            ELSIF fbReceive.nRecBytes > 0 THEN
                nRxCount := nRxCount + fbReceive.nRecBytes;
                IF nRxCount >= 9 THEN
                    nExpectedFrame := 9 + BYTE_TO_UDINT(aRx[7]) + BYTE_TO_UDINT(aRx[8]) * 256;
                    IF (nExpectedFrame < 11) OR (nExpectedFrame > SIZEOF(aRx)) THEN
                        bError := TRUE; nErrorID := 16#E104;
                        stSession.bConnected := FALSE;
                        bBusy := FALSE; nState := 0;
                    ELSIF nRxCount >= nExpectedFrame THEN
                        IF (aRx[0] <> 16#D0) OR (aRx[1] <> 16#00) THEN
                            bError := TRUE; nErrorID := 16#E105;
                            stSession.bConnected := FALSE;
                        ELSE
                            nEndCode := BYTE_TO_UINT(aRx[9]) + BYTE_TO_UINT(aRx[10]) * 256;
                            IF nEndCode <> 0 THEN
                                bError := TRUE; nErrorID := nEndCode;
                            ELSIF (bBitAccess AND (nExpectedFrame < 11 + ((UINT_TO_UDINT(nPoints) + 1) / 2)))
                                 OR ((NOT bBitAccess) AND (nExpectedFrame < 11 + UINT_TO_UDINT(nPoints) * 2)) THEN
                                bError := TRUE; nErrorID := 16#E107;
                                stSession.bConnected := FALSE;
                            ELSE
                                IF bBitAccess THEN
                                    pDestBit := pData;
                                    FOR nIdx := 0 TO (UINT_TO_UDINT(nPoints) - 1) DO
                                        IF (nIdx MOD 2) = 0 THEN
                                            pDestBit[nIdx] := ((aRx[11 + (nIdx / 2)] AND 16#10) <> 0);
                                        ELSE
                                            pDestBit[nIdx] := ((aRx[11 + (nIdx / 2)] AND 16#01) <> 0);
                                        END_IF;
                                    END_FOR;
                                ELSE
                                    pDestByte := pData;
                                    nCopyBytes := UINT_TO_UDINT(nPoints) * 2;
                                    FOR nIdx := 0 TO (nCopyBytes - 1) DO
                                        pDestByte[nIdx] := aRx[11 + nIdx];
                                    END_FOR;
                                END_IF;
                                bDone := TRUE;
                            END_IF;
                        END_IF;
                        bBusy := FALSE; nState := 0;
                    ELSE
                        nState := 20; // Fragment received; wait for rest of frame
                    END_IF;
                ELSE
                    nState := 20; // Header itself is fragmented
                END_IF;

            ELSIF tonTimeout.Q THEN
                // Quá 2 giây không có phản hồi
                bError   := TRUE;
                nErrorID := 16#E103; // Timeout chờ response
                stSession.bConnected := FALSE;
                bBusy    := FALSE;
                nState   := 0;

            ELSE
                // Chưa có dữ liệu về trong scan này -> Kích đọc tiếp ở scan sau
                nState := 20;
            END_IF;
        END_IF;

END_CASE;

// Cập nhật trạng thái bận vào session dùng chung
// Only the FB that acquired the socket lock may release it.
IF bBusy THEN
    stSession.bBusy := TRUE;
ELSIF bOwnsSession THEN
    stSession.bBusy := FALSE;
    bOwnsSession := FALSE;
END_IF;

END_FUNCTION_BLOCK

// ---- POUs/FB_MelsecDebugXY4Pt.TcPOU
FUNCTION_BLOCK FB_MelsecDebugXY4Pt
VAR_INPUT
    bExecute          : BOOL := FALSE; // Rising edge for ONE 4-point DATA-ONLY test
    bPermit           : BOOL := FALSE; // Maintenance gate, OFF by default
    bMachineStopped   : BOOL := FALSE; // Axis, encoder and gantry are stationary
    bPublisherIdle    : BOOL := FALSE; // All live motion publishers inhibited
    bAbort            : BOOL := FALSE; // Cancel the data-only sequence
    rCenterX_mm       : LREAL := 50.0;
    rCenterY_mm       : LREAL := 85.0;
    rAngleDeg         : LREAL := 0.0;
    rLength_mm        : LREAL := 40.0;
    rWidth_mm         : LREAL := 40.0;
    tHold             : TIME := T#10S; // GX Works2 observation pause, NOT motion acknowledgment
END_VAR
VAR_IN_OUT
    stSession         : ST_MelsecSession; // Same owned socket as all other TwinCAT FBs
END_VAR
VAR_OUTPUT
    bBusy             : BOOL;
    bDone             : BOOL;       // Four XY frames READ BACK; NOT robot motion completion
    bError            : BOOL;
    nErrorCode        : INT;
    nCommErrorID      : UDINT;
    nState            : INT := 0;
    nCurrentVertex    : INT;        // 1..4, stays at 4 after success
    nPassedVertices   : INT;
    nWriteX           : DINT;
    nWriteY           : DINT;
    nReadX            : DINT;
    nReadY            : DINT;
    nReadVertex       : UINT;
    bLastReadbackOK   : BOOL;
    bAllMotionBitsLow : BOOL;
    bOriginalRestored : BOOL; // Original XY/index restored after all four hold windows
END_VAR
VAR
    fbStart           : R_TRIG;
    fbWrite           : FB_MelsecWrite;
    fbRead            : FB_MelsecRead;
    tonHold           : TON;
    aCorners          : ARRAY[1..4] OF ST_Point2D;
    rAngleRad         : LREAL;
    rC                : LREAL;
    rS                : LREAL;
    rHL               : LREAL;
    rHW               : LREAL;
    aXYWrite          : ARRAY[0..1] OF DINT;
    aXYRead           : ARRAY[0..1] OF DINT;
    nIndexWrite       : UINT;
    nIndexRead        : UINT;
    aOriginalXY       : ARRAY[0..1] OF DINT;
    nOriginalIndex    : UINT;
    bNeedSnapshot     : BOOL;
    bRestoring        : BOOL;
    aStartAck         : ARRAY[0..1] OF BOOL; // M1000 M1001
    aRobotFlags       : ARRAY[0..3] OF BOOL; // M102, M103, M104, M105
    nPlcFsmState      : DINT;               // D200/D201
    bWriteReq         : BOOL;
    bReadReq          : BOOL;
    eReadDevice       : E_MelsecDevice;
    nReadAddress      : UDINT;
    nReadPoints       : UINT;
    bReadBitMode      : BOOL;
    pReadData         : PVOID;
    nReadDataSize     : UDINT;
    nWriteAddress     : UDINT;
    nWritePoints      : UINT;
    pWriteData        : PVOID;
    nWriteDataSize    : UDINT;
END_VAR

// Diagnostic mode NEVER writes M1000 or any PLC bit, never touches Z.
// Only D100..D103 (2x DINT XY) and D114 (UINT vertex) are ever written.
// Explicit machine-stopped conditions are checked on EVERY scan.
fbStart(CLK := bExecute);
tonHold(IN := (nState = 20), PT := tHold);

bReadReq := FALSE;
bWriteReq := FALSE;

IF (nState <> 0) AND (nState <> 99) AND (NOT bPermit OR NOT bMachineStopped OR
    NOT bPublisherIdle OR bAbort OR NOT stSession.bConnected) THEN
    bError := TRUE;
    nErrorCode := 901; // Lost permit, motion interlock, or TCP
    nState := 99;
END_IF;

CASE nState OF
    0: // IDLE - no automatic restart
        bBusy := FALSE;
        IF fbStart.Q THEN
            bDone := FALSE;
            bError := FALSE;
            bLastReadbackOK := FALSE;
            bAllMotionBitsLow := FALSE;
            nPassedVertices := 0;
            nCurrentVertex := 0;
            bNeedSnapshot := TRUE;
            bRestoring := FALSE;
            bOriginalRestored := FALSE;
            nErrorCode := 0;
            nCommErrorID := 0;
            IF NOT bPermit OR NOT bMachineStopped OR NOT bPublisherIdle
                OR bAbort OR NOT stSession.bConnected OR stSession.bBusy THEN
                bError := TRUE; nErrorCode := 901;
            ELSIF (rLength_mm <= 0.0) OR (rWidth_mm <= 0.0)
                OR (rLength_mm > 100.0) OR (rWidth_mm > 100.0)
                OR (tHold < T#2S) OR (tHold > T#60S) THEN
                bError := TRUE; nErrorCode := 902;
            ELSE
                rAngleRad := rAngleDeg * 3.141592653589793 / 180.0;
                rC := COS(rAngleRad);
                rS := SIN(rAngleRad);
                rHL := rLength_mm / 2.0;
                rHW := rWidth_mm / 2.0;

                aCorners[1].X := rCenterX_mm + rHL * rC - rHW * rS;
                aCorners[1].Y := rCenterY_mm + rHL * rS + rHW * rC;
                aCorners[2].X := rCenterX_mm - rHL * rC - rHW * rS;
                aCorners[2].Y := rCenterY_mm - rHL * rS + rHW * rC;
                aCorners[3].X := rCenterX_mm - rHL * rC + rHW * rS;
                aCorners[3].Y := rCenterY_mm - rHL * rS - rHW * rC;
                aCorners[4].X := rCenterX_mm + rHL * rC + rHW * rS;
                aCorners[4].Y := rCenterY_mm + rHL * rS - rHW * rC;

                nCurrentVertex := 1;
                bBusy := TRUE;
                nState := 1;
            END_IF;
        END_IF;

    // Recheck Mitsubishi handshake before EVERY vertex (read-only).
    1:
        eReadDevice := DEV_M; nReadAddress := 1000; nReadPoints := 2;
        bReadBitMode := TRUE;
        pReadData := ADR(aStartAck); nReadDataSize := SIZEOF(aStartAck);
        bReadReq := TRUE;
        nState := 2;

    2:
        IF fbRead.bDone THEN
            IF aStartAck[0] OR aStartAck[1] THEN
                bError := TRUE; nErrorCode := 903; nState := 99;
            ELSE
                nState := 3;
            END_IF;
        ELSIF fbRead.bError THEN
            bError := TRUE; nErrorCode := 910; nCommErrorID := fbRead.nErrorID; nState := 99;
        END_IF;

    3:
        eReadDevice := DEV_M; nReadAddress := 102; nReadPoints := 4;
        bReadBitMode := TRUE;
        pReadData := ADR(aRobotFlags); nReadDataSize := SIZEOF(aRobotFlags);
        bReadReq := TRUE;
        nState := 4;

    4:
        IF fbRead.bDone THEN
            IF aRobotFlags[0] OR aRobotFlags[1] OR aRobotFlags[2] OR aRobotFlags[3] THEN
                bError := TRUE; nErrorCode := 904; nState := 99;
            ELSE
                nState := 5;
            END_IF;
        ELSIF fbRead.bError THEN
            bError := TRUE; nErrorCode := 911; nCommErrorID := fbRead.nErrorID; nState := 99;
        END_IF;

    5:
        eReadDevice := DEV_D; nReadAddress := 200; nReadPoints := 2;
        bReadBitMode := FALSE;
        pReadData := ADR(nPlcFsmState); nReadDataSize := SIZEOF(nPlcFsmState);
        bReadReq := TRUE;
        nState := 6;

    6:
        IF fbRead.bDone THEN
            IF nPlcFsmState <> 0 THEN
                bError := TRUE; nErrorCode := 905; nState := 99;
            ELSE
                bAllMotionBitsLow := TRUE;
                IF bRestoring THEN
                    nState := 30;
                ELSIF bNeedSnapshot THEN
                    nState := 7;
                ELSE
                    nState := 10;
                END_IF;
            END_IF;
        ELSIF fbRead.bError THEN
            bError := TRUE; nErrorCode := 912; nCommErrorID := fbRead.nErrorID; nState := 99;
        END_IF;

    7: // Snapshot original XY before any data-only write
        eReadDevice := DEV_D; nReadAddress := 100; nReadPoints := 4;
        bReadBitMode := FALSE;
        pReadData := ADR(aOriginalXY); nReadDataSize := SIZEOF(aOriginalXY);
        bReadReq := TRUE;
        nState := 8;

    8:
        IF fbRead.bDone THEN
            nState := 9;
        ELSIF fbRead.bError THEN
            bError := TRUE; nErrorCode := 918; nCommErrorID := fbRead.nErrorID; nState := 99;
        END_IF;

    9:
        eReadDevice := DEV_D; nReadAddress := 114; nReadPoints := 1;
        bReadBitMode := FALSE;
        pReadData := ADR(nOriginalIndex); nReadDataSize := SIZEOF(nOriginalIndex);
        bReadReq := TRUE;
        nState := 91;

    91:
        IF fbRead.bDone THEN
            bNeedSnapshot := FALSE;
            nState := 10;
        ELSIF fbRead.bError THEN
            bError := TRUE; nErrorCode := 919; nCommErrorID := fbRead.nErrorID; nState := 99;
        END_IF;

    10: // Data-only: two DINTs. Deliberately no Z/speed write.
        IF (nCurrentVertex < 1) OR (nCurrentVertex > 4) OR
            (aCorners[nCurrentVertex].X < 5.0) OR
            (aCorners[nCurrentVertex].X > 170.0) OR
            (aCorners[nCurrentVertex].Y < 5.0) OR
            (aCorners[nCurrentVertex].Y > 165.0) THEN
            bError := TRUE; nErrorCode := 906; nState := 99;
        ELSE
            nWriteX := LREAL_TO_DINT(aCorners[nCurrentVertex].X * 10000.0);
            nWriteY := LREAL_TO_DINT(aCorners[nCurrentVertex].Y * 10000.0);
            aXYWrite[0] := nWriteX;
            aXYWrite[1] := nWriteY;
            nIndexWrite := INT_TO_UINT(nCurrentVertex);
            nWriteAddress := 100; nWritePoints := 4;
            pWriteData := ADR(aXYWrite); nWriteDataSize := SIZEOF(aXYWrite);
            bLastReadbackOK := FALSE;
            bWriteReq := TRUE;
            nState := 11;
        END_IF;

    11:
        IF fbWrite.bDone THEN
            nState := 12;
        ELSIF fbWrite.bError THEN
            bError := TRUE; nErrorCode := 913; nCommErrorID := fbWrite.nErrorID; nState := 99;
        END_IF;

    12: // Different rising edge for D114
        nWriteAddress := 114; nWritePoints := 1;
        pWriteData := ADR(nIndexWrite); nWriteDataSize := SIZEOF(nIndexWrite);
        bWriteReq := TRUE;
        nState := 13;

    13:
        IF fbWrite.bDone THEN
            nState := 14;
        ELSIF fbWrite.bError THEN
            bError := TRUE; nErrorCode := 914; nCommErrorID := fbWrite.nErrorID; nState := 99;
        END_IF;

    14:
        eReadDevice := DEV_D; nReadAddress := 100; nReadPoints := 4;
        bReadBitMode := FALSE;
        pReadData := ADR(aXYRead); nReadDataSize := SIZEOF(aXYRead);
        bReadReq := TRUE;
        nState := 15;

    15:
        IF fbRead.bDone THEN
            nState := 16;
        ELSIF fbRead.bError THEN
            bError := TRUE; nErrorCode := 915; nCommErrorID := fbRead.nErrorID; nState := 99;
        END_IF;

    16:
        eReadDevice := DEV_D; nReadAddress := 114; nReadPoints := 1;
        bReadBitMode := FALSE;
        pReadData := ADR(nIndexRead); nReadDataSize := SIZEOF(nIndexRead);
        bReadReq := TRUE;
        nState := 17;

    17:
        IF fbRead.bDone THEN
            nReadX := aXYRead[0];
            nReadY := aXYRead[1];
            nReadVertex := nIndexRead;
            bLastReadbackOK := (nReadX = nWriteX) AND (nReadY = nWriteY)
                               AND (nReadVertex = nIndexWrite);
            IF bLastReadbackOK THEN
                nPassedVertices := nPassedVertices + 1;
                nState := 20; // Hold for operator GX Works2 observation
            ELSE
                bError := TRUE; nErrorCode := 916; nState := 99;
            END_IF;
        ELSIF fbRead.bError THEN
            bError := TRUE; nErrorCode := 917; nCommErrorID := fbRead.nErrorID; nState := 99;
        END_IF;

    20: // Observation timer. Never mislabel elapsed time as QD75 motion ACK.
        IF tonHold.Q THEN
            IF nCurrentVertex >= 4 THEN
                bRestoring := TRUE;
                bAllMotionBitsLow := FALSE;
                nState := 1; // Recheck M1000/ACK/BUSY/FSM before restoring original packet
            ELSE
                nCurrentVertex := nCurrentVertex + 1;
                bAllMotionBitsLow := FALSE;
                nState := 1;
            END_IF;
        END_IF;

    30: // Restore original XY, then original index: never leave stale debug target
        nWriteAddress := 100; nWritePoints := 4;
        pWriteData := ADR(aOriginalXY); nWriteDataSize := SIZEOF(aOriginalXY);
        bWriteReq := TRUE;
        nState := 31;

    31:
        IF fbWrite.bDone THEN
            nState := 32;
        ELSIF fbWrite.bError THEN
            bError := TRUE; nErrorCode := 920; nCommErrorID := fbWrite.nErrorID; nState := 99;
        END_IF;

    32:
        nWriteAddress := 114; nWritePoints := 1;
        pWriteData := ADR(nOriginalIndex); nWriteDataSize := SIZEOF(nOriginalIndex);
        bWriteReq := TRUE;
        nState := 33;

    33:
        IF fbWrite.bDone THEN
            nState := 34;
        ELSIF fbWrite.bError THEN
            bError := TRUE; nErrorCode := 921; nCommErrorID := fbWrite.nErrorID; nState := 99;
        END_IF;

    34:
        eReadDevice := DEV_D; nReadAddress := 100; nReadPoints := 4;
        bReadBitMode := FALSE;
        pReadData := ADR(aXYRead); nReadDataSize := SIZEOF(aXYRead);
        bReadReq := TRUE;
        nState := 35;

    35:
        IF fbRead.bDone THEN
            nState := 36;
        ELSIF fbRead.bError THEN
            bError := TRUE; nErrorCode := 922; nCommErrorID := fbRead.nErrorID; nState := 99;
        END_IF;

    36:
        eReadDevice := DEV_D; nReadAddress := 114; nReadPoints := 1;
        bReadBitMode := FALSE;
        pReadData := ADR(nIndexRead); nReadDataSize := SIZEOF(nIndexRead);
        bReadReq := TRUE;
        nState := 37;

    37:
        IF fbRead.bDone THEN
            bOriginalRestored := (aXYRead[0] = aOriginalXY[0]) AND
                (aXYRead[1] = aOriginalXY[1]) AND (nIndexRead = nOriginalIndex);
            IF bOriginalRestored THEN
                bBusy := FALSE;
                bDone := TRUE; // All 4 readbacks AND full restore confirmed
                nState := 0;
            ELSE
                bError := TRUE; nErrorCode := 923; nState := 99;
            END_IF;
        ELSIF fbRead.bError THEN
            bError := TRUE; nErrorCode := 924; nCommErrorID := fbRead.nErrorID; nState := 99;
        END_IF;

    99: // Latched diagnostic failure. NO reset command sent to the PLC.
        bBusy := FALSE;
        bDone := FALSE;
        bReadReq := FALSE;
        bWriteReq := FALSE;
        IF NOT bExecute AND NOT bPermit AND NOT fbRead.bBusy AND NOT fbWrite.bBusy THEN
            nState := 0;
        END_IF;
END_CASE;

// READS may access only M1000,M1001,M102..M105,D200..D201,D100..D103,D114.
// WRITES are strictly limited to D100..D103 and D114, never M, Z or QD75.
fbWrite(
    stSession := stSession, bExecute := bWriteReq,
    eDevice := DEV_D, nStartAddr := nWriteAddress,
    nPoints := nWritePoints, bBitAccess := FALSE,
    pData := pWriteData, nDataSize := nWriteDataSize
);
fbRead(
    stSession := stSession, bExecute := bReadReq,
    eDevice := eReadDevice, nStartAddr := nReadAddress,
    nPoints := nReadPoints, bBitAccess := bReadBitMode,
    pData := pReadData, nDataSize := nReadDataSize
);

END_FUNCTION_BLOCK

// ---- POUs/FB_UpstreamCameraTracking4Pt.TcPOU
FUNCTION_BLOCK FB_UpstreamCameraTracking4Pt
VAR_INPUT
    bReset               : BOOL;
    bCameraResult        : BOOL;  // Single rising edge: camera provides center and angle ONLY
    bAcceptCamera        : BOOL;
    bCalibrationConfirmed: BOOL;  // NEVER assume Camera and Robot coordinates coincide
    bExposureEncoderValid : BOOL; // Capture encoder synchronized with IMAGE EXPOSURE, not processing result
    rEncoderAtExposure_mm : LREAL; // Encoder latched by TwinCAT when camera takes the image
    rCameraCenterX_mm    : LREAL; // Already calibrated from pixels into millimeters
    rCameraCenterY_mm    : LREAL;
    rCameraAngleDeg      : LREAL;
    rCameraToWorkStart_mm : LREAL; // USER INPUT after calibration: Camera trigger station to ROBOT X=0, positive mm
    rCameraToRobotX_mm   : LREAL; // Fine X calibration correction only; NOT the Camera->Robot distance
    rCameraToRobotY_mm   : LREAL;
    rCameraToRobotYawDeg : LREAL; // Calibrated camera-to-robot axis angle
    rEncoderTotalDist_mm : LREAL; // Continuous integrated encoder distance, not 16-bit count
    rLength_mm           : LREAL := 40.0;
    rWidth_mm            : LREAL := 40.0;
    rRobotXMin_mm        : LREAL := 0.0;
    rRobotXMax_mm        : LREAL := 180.0;
    rRobotYMin_mm        : LREAL := 0.0;
    rRobotYMax_mm        : LREAL := 170.0;
END_VAR
VAR_OUTPUT
    bCaptured            : BOOL; // Product retained while travelling FROM camera to robot
    bInRobotWorkspace    : BOOL; // At least one corner in workspace (diagnostic only)
    bAllCornersPastRobot : BOOL;
    bCalibrationMissing  : BOOL;
    nCaptureCount        : UDINT;
    nRejectedCount       : UDINT;
    nErrorCode           : INT;
    rEncoderAtCapture_mm : LREAL;
    rEncoderTravel_mm    : LREAL;
    rCenterAtCaptureX_mm : LREAL; // Robot reference frame at camera trigger time
    rCenterAtCaptureY_mm : LREAL;
    rThetaRobotDeg       : LREAL;
    rCenterNowX_mm       : LREAL; // Current center position in robot frame, negative upstream
    rCenterNowY_mm       : LREAL;
    rToRobotWorkStart_mm : LREAL; // Positive while center still upstream; 0 once X>=0
    aCornerAtCamera      : ARRAY[1..4] OF ST_Point2D;
    aCornerNow           : ARRAY[1..4] OF ST_Point2D;
END_VAR
VAR
    fbCameraEdge         : R_TRIG;
    bFirstScan           : BOOL := TRUE;
    bStartupReset        : BOOL;
    rFrameRad            : LREAL;
    rPhiC                : LREAL;
    rPhiS                : LREAL;
    rThetaRad            : LREAL;
    rC                  : LREAL;
    rS                  : LREAL;
    rHx                 : LREAL;
    rHy                 : LREAL;
    aLocalX             : ARRAY[1..4] OF LREAL;
    aLocalY             : ARRAY[1..4] OF LREAL;
    i                    : INT;
END_VAR

fbCameraEdge(CLK := bCameraResult);
bCalibrationMissing := NOT bCalibrationConfirmed
    OR (rCameraToWorkStart_mm <= 0.0) OR (rCameraToWorkStart_mm > 100000.0);

// Startup: zero LOGICAL state only. Do NOT reset physical encoder/servo.
// bReset can also be issued deliberately while offline/idle.
bStartupReset := bFirstScan OR bReset;
IF bStartupReset THEN
    bFirstScan := FALSE;
    bCaptured := FALSE;
    bInRobotWorkspace := FALSE;
    bAllCornersPastRobot := FALSE;
    nCaptureCount := 0;
    nRejectedCount := 0;
    nErrorCode := 0;
    rEncoderAtCapture_mm := 0.0;
    rEncoderTravel_mm := 0.0;
    rCenterAtCaptureX_mm := 0.0;
    rCenterAtCaptureY_mm := 0.0;
    rCenterNowX_mm := 0.0;
    rCenterNowY_mm := 0.0;
    rToRobotWorkStart_mm := 0.0;
    rThetaRobotDeg := 0.0;
    FOR i := 1 TO 4 DO
        aCornerAtCamera[i].X := 0.0;
        aCornerAtCamera[i].Y := 0.0;
        aCornerNow[i].X := 0.0;
        aCornerNow[i].Y := 0.0;
    END_FOR;
END_IF;

IF fbCameraEdge.Q AND NOT bStartupReset THEN
    IF bCalibrationMissing OR NOT bAcceptCamera OR bCaptured OR NOT bExposureEncoderValid THEN
        nRejectedCount := nRejectedCount + 1;
        nErrorCode := 101; // Invalid calibration or previously tracked product
    ELSIF (rLength_mm <= 0.0) OR (rWidth_mm <= 0.0)
       OR (rLength_mm > 100.0) OR (rWidth_mm > 100.0)
       OR (ABS(rCameraCenterX_mm) > 100000.0)
       OR (ABS(rCameraCenterY_mm) > 100000.0) THEN
        nRejectedCount := nRejectedCount + 1;
        nErrorCode := 102;
    ELSE
        // Frame transform: coordinates in camera physical mm, to robot mm.
        // Pixel -> mm calibration must happen BEFORE this FB.
        rFrameRad := rCameraToRobotYawDeg * 3.141592653589793 / 180.0;
        rPhiC := COS(rFrameRad);
        rPhiS := SIN(rFrameRad);
        rCenterAtCaptureX_mm :=
            -rCameraToWorkStart_mm + rCameraToRobotX_mm
            + rCameraCenterX_mm * rPhiC - rCameraCenterY_mm * rPhiS;
        rCenterAtCaptureY_mm :=
            rCameraToRobotY_mm + rCameraCenterX_mm * rPhiS + rCameraCenterY_mm * rPhiC;
        rThetaRobotDeg := rCameraAngleDeg + rCameraToRobotYawDeg;
        rThetaRad := rThetaRobotDeg * 3.141592653589793 / 180.0;
        rC := COS(rThetaRad);
        rS := SIN(rThetaRad);
        rHx := rLength_mm / 2.0;
        rHy := rWidth_mm / 2.0;

        aLocalX[1] := rHx;  aLocalY[1] := rHy;
        aLocalX[2] := -rHx; aLocalY[2] := rHy;
        aLocalX[3] := -rHx; aLocalY[3] := -rHy;
        aLocalX[4] := rHx;  aLocalY[4] := -rHy;
        FOR i := 1 TO 4 DO
            aCornerAtCamera[i].X := rCenterAtCaptureX_mm +
                aLocalX[i] * rC - aLocalY[i] * rS;
            aCornerAtCamera[i].Y := rCenterAtCaptureY_mm +
                aLocalX[i] * rS + aLocalY[i] * rC;
            aCornerNow[i] := aCornerAtCamera[i];
        END_FOR;
        rEncoderAtCapture_mm := rEncoderAtExposure_mm;
        rEncoderTravel_mm := 0.0;
        bCaptured := TRUE;
        bAllCornersPastRobot := FALSE;
        nCaptureCount := nCaptureCount + 1;
        nErrorCode := 0;
    END_IF;
END_IF;

IF bCaptured THEN
    rEncoderTravel_mm := rEncoderTotalDist_mm - rEncoderAtCapture_mm;
    rCenterNowX_mm := rCenterAtCaptureX_mm + rEncoderTravel_mm;
    rCenterNowY_mm := rCenterAtCaptureY_mm;
    IF rCenterNowX_mm < 0.0 THEN
        rToRobotWorkStart_mm := -rCenterNowX_mm;
    ELSE
        rToRobotWorkStart_mm := 0.0;
    END_IF;
    bInRobotWorkspace := FALSE;
    bAllCornersPastRobot := TRUE;
    FOR i := 1 TO 4 DO
        aCornerNow[i].X := aCornerAtCamera[i].X + rEncoderTravel_mm;
        aCornerNow[i].Y := aCornerAtCamera[i].Y;
        IF (aCornerNow[i].X >= rRobotXMin_mm)
           AND (aCornerNow[i].X <= rRobotXMax_mm)
           AND (aCornerNow[i].Y >= rRobotYMin_mm)
           AND (aCornerNow[i].Y <= rRobotYMax_mm) THEN
            bInRobotWorkspace := TRUE;
        END_IF;
        IF aCornerNow[i].X <= rRobotXMax_mm THEN
            bAllCornersPastRobot := FALSE;
        END_IF;
    END_FOR;
    // Unlike the old FB, upstream negative-X locations remain valid!
    IF bAllCornersPastRobot THEN
        bCaptured := FALSE;
        nErrorCode := 103; // Product exited workspace
    END_IF;
END_IF;

END_FUNCTION_BLOCK

// ---- POUs/FB_CameraProductQueue.TcPOU
FUNCTION_BLOCK FB_CameraProductQueue
VAR_INPUT
    bReset                  : BOOL;
    bLiveExposure           : BOOL; // physical image-exposure signal (NOT camera result)
    bLiveResult             : BOOL; // result contains calibrated X/Y mm + angle
    bLiveBridgeVerified     : BOOL; // FALSE until real camera driver audited
    bCalibrationConfirmed   : BOOL; // FALSE until camera -> robot calibration audited

    // BENCH SIMULATION ONLY: not linked to robot publisher / M1000
    bSimMode                : BOOL;
    bSimExposure            : BOOL;
    bSimResult              : BOOL;
    bSimCompleteHead        : BOOL;

    rCenterX_mm             : LREAL;
    rCenterY_mm             : LREAL;
    rAngle_deg              : LREAL;
    rCameraToWorkStart_mm   : LREAL; // calibrated positive distance to ROBOT X=0
    rCameraFineOffsetX_mm   : LREAL;
    rCameraOffsetY_mm       : LREAL;
    rCameraYaw_deg          : LREAL;
    rLength_mm              : LREAL := 40.0;
    rWidth_mm               : LREAL := 40.0;
    rEncoderTotalDist_mm    : LREAL; // integrated distance, NOT 16-bit raw pulse
    rConveyorSpeed_mm_s     : LREAL;
    rXMin_mm                : LREAL := 0.0;
    rXMax_mm                : LREAL := 180.0;
    rYMin_mm                : LREAL := 0.0;
    rYMax_mm                : LREAL := 170.0;
    rMinCycleBudget_s       : LREAL := 1.2;  // planning estimate, NOT validated robot duration
    rFlyTime_s              : LREAL := 0.12;
    rSyncTime_s             : LREAL := 0.06;
END_VAR
VAR_OUTPUT
    aQueue                  : ARRAY[1..8] OF ST_QueuedCameraProduct;
    nQueueCount             : INT;
    nHeadIndex              : INT := 1;
    nTailIndex              : INT := 1;
    nHeadProductID          : UDINT;
    nHeadState              : INT;
    nLastAcceptedProductID  : UDINT;
    nAccepted               : UDINT;
    nRejected               : UDINT;
    nMissed                 : UDINT;
    nSimCompleted           : UDINT; // BENCH simulator ONLY, not robot done
    nExposureOverruns       : UDINT;
    nErrorCode              : INT;
    bInputFault             : BOOL; // latched until reset
    bPendingExposure        : BOOL;
    bQueueFull              : BOOL;
    bHeadValid              : BOOL;
    bHeadAllInside          : BOOL;
    bHeadForecastOK         : BOOL; // geometry/timing estimate ONLY, no motion authorization
    rHeadTravel_mm          : LREAL;
    rHeadToWorkStart_mm     : LREAL;
    rHeadCenterX_mm         : LREAL;
    rHeadCenterY_mm         : LREAL;
    aHeadCornerNow          : ARRAY[1..4] OF ST_Point2D;
END_VAR
VAR
    fbExposureEdge          : R_TRIG;
    fbResultEdge            : R_TRIG;
    fbSimDoneEdge           : R_TRIG;
    tonResultTTL            : TON;
    bFirstScan              : BOOL := TRUE;
    rPendingEncoder_mm      : LREAL;
    rYawRad                 : LREAL;
    rThetaRad               : LREAL;
    rCosYaw                 : LREAL;
    rSinYaw                 : LREAL;
    rCosTheta               : LREAL;
    rSinTheta               : LREAL;
    rHalfL                  : LREAL;
    rHalfW                  : LREAL;
    rLocalX                 : LREAL;
    rLocalY                 : LREAL;
    rCenterRobotX           : LREAL;
    rCenterRobotY           : LREAL;
    rForecastMotion_mm      : LREAL;
    bOut                    : BOOL;
    i                       : INT;
    j                       : INT;
    nSlot                   : INT;
END_VAR

// STAGED DATA-ONLY FIFO: no MC writes, no M1000, no QD75 and no servo output.
// A single unmatched exposure is allowed at a time because the camera has
// not yet provided frame IDs. Overlapping exposures cause a latched fault.
fbExposureEdge(CLK := (bLiveExposure AND bLiveBridgeVerified AND NOT bSimMode)
                        OR (bSimExposure AND bSimMode));
fbResultEdge(CLK := (bLiveResult AND bLiveBridgeVerified AND NOT bSimMode)
                      OR (bSimResult AND bSimMode));
fbSimDoneEdge(CLK := bSimCompleteHead AND bSimMode);
tonResultTTL(IN := bPendingExposure, PT := T#5S);

IF bFirstScan OR bReset THEN
    bFirstScan := FALSE;
    nQueueCount := 0;
    nHeadIndex := 1;
    nTailIndex := 1;
    nHeadProductID := 0;
    nHeadState := 0;
    nLastAcceptedProductID := 0;
    nAccepted := 0;
    nRejected := 0;
    nMissed := 0;
    nSimCompleted := 0;
    nExposureOverruns := 0;
    nErrorCode := 0;
    bInputFault := FALSE;
    bPendingExposure := FALSE;
    bQueueFull := FALSE;
    bHeadValid := FALSE;
    bHeadAllInside := FALSE;
    bHeadForecastOK := FALSE;
    rPendingEncoder_mm := 0.0;
    rHeadTravel_mm := 0.0;
    rHeadToWorkStart_mm := 0.0;
    rHeadCenterX_mm := 0.0;
    rHeadCenterY_mm := 0.0;
    FOR i := 1 TO 8 DO
        aQueue[i].bValid := FALSE;
        aQueue[i].nState := 0;
        aQueue[i].nProductID := 0;
        aQueue[i].bAllCornersInside := FALSE;
        aQueue[i].bForecastWindowOK := FALSE;
        aQueue[i].rEncoderAtExposure_mm := 0.0;
        aQueue[i].rCenterAtExposureX_mm := 0.0;
        aQueue[i].rCenterAtExposureY_mm := 0.0;
        aQueue[i].rThetaRobot_deg := 0.0;
        aQueue[i].rTravel_mm := 0.0;
        aQueue[i].rCenterNowX_mm := 0.0;
        aQueue[i].rCenterNowY_mm := 0.0;
        FOR j := 1 TO 4 DO
            aQueue[i].aCornerBase[j].X := 0.0;
            aQueue[i].aCornerBase[j].Y := 0.0;
            aQueue[i].aCornerNow[j].X := 0.0;
            aQueue[i].aCornerNow[j].Y := 0.0;
        END_FOR;
    END_FOR;
END_IF;

IF NOT bReset THEN
    IF bPendingExposure AND tonResultTTL.Q THEN
        bPendingExposure := FALSE;
        bInputFault := TRUE;
        nErrorCode := 110; // Camera processing result exceeded 5 seconds
        nRejected := nRejected + 1;
    END_IF;

    IF fbExposureEdge.Q THEN
        IF bInputFault OR bPendingExposure THEN
            bInputFault := TRUE; // no frame-ID: cannot pair overlapping images
            bPendingExposure := FALSE;
            nExposureOverruns := nExposureOverruns + 1;
            nErrorCode := 111;
        ELSIF (rCameraToWorkStart_mm <= 0.0)
            OR (rCameraToWorkStart_mm > 100000.0)
            OR (NOT bCalibrationConfirmed AND NOT bSimMode) THEN
            nRejected := nRejected + 1;
            nErrorCode := 112; // no physically verified calibration
        ELSE
            rPendingEncoder_mm := rEncoderTotalDist_mm;
            bPendingExposure := TRUE;
        END_IF;
    END_IF;

    IF fbResultEdge.Q THEN
        IF bInputFault OR NOT bPendingExposure THEN
            nRejected := nRejected + 1;
            nErrorCode := 113; // result without matching exposure
        ELSIF (rLength_mm <= 0.0) OR (rWidth_mm <= 0.0)
            OR (rLength_mm > 100.0) OR (rWidth_mm > 100.0)
            OR (ABS(rCenterX_mm) > 100000.0)
            OR (ABS(rCenterY_mm) > 100000.0)
            OR (ABS(rAngle_deg) > 3600.0) THEN
            nRejected := nRejected + 1;
            nErrorCode := 114;
            bPendingExposure := FALSE;
        ELSIF nQueueCount >= 8 THEN
            nRejected := nRejected + 1;
            nErrorCode := 115; // full; never overwrite a live product
            bQueueFull := TRUE;
            bPendingExposure := FALSE;
        ELSE
            nSlot := nTailIndex;
            rYawRad := rCameraYaw_deg * 3.141592653589793 / 180.0;
            rCosYaw := COS(rYawRad);
            rSinYaw := SIN(rYawRad);
            rCenterRobotX := -rCameraToWorkStart_mm + rCameraFineOffsetX_mm
                + rCenterX_mm * rCosYaw - rCenterY_mm * rSinYaw;
            rCenterRobotY := rCameraOffsetY_mm
                + rCenterX_mm * rSinYaw + rCenterY_mm * rCosYaw;
            rThetaRad := (rAngle_deg + rCameraYaw_deg)
                * 3.141592653589793 / 180.0;
            rCosTheta := COS(rThetaRad);
            rSinTheta := SIN(rThetaRad);
            rHalfL := rLength_mm / 2.0;
            rHalfW := rWidth_mm / 2.0;
            aQueue[nSlot].bValid := TRUE;
            aQueue[nSlot].nState := 1; // WAIT_ROBOT
            nLastAcceptedProductID := nLastAcceptedProductID + 1;
            aQueue[nSlot].nProductID := nLastAcceptedProductID;
            aQueue[nSlot].rEncoderAtExposure_mm := rPendingEncoder_mm;
            aQueue[nSlot].rCenterAtExposureX_mm := rCenterRobotX;
            aQueue[nSlot].rCenterAtExposureY_mm := rCenterRobotY;
            aQueue[nSlot].rThetaRobot_deg := rAngle_deg + rCameraYaw_deg;
            aQueue[nSlot].rTravel_mm := 0.0;
            aQueue[nSlot].rCenterNowX_mm := rCenterRobotX;
            aQueue[nSlot].rCenterNowY_mm := rCenterRobotY;
            FOR j := 1 TO 4 DO
                CASE j OF
                    1: rLocalX := rHalfL;  rLocalY := rHalfW;
                    2: rLocalX := -rHalfL; rLocalY := rHalfW;
                    3: rLocalX := -rHalfL; rLocalY := -rHalfW;
                    4: rLocalX := rHalfL;  rLocalY := -rHalfW;
                END_CASE;
                aQueue[nSlot].aCornerBase[j].X := rCenterRobotX
                    + rLocalX * rCosTheta - rLocalY * rSinTheta;
                aQueue[nSlot].aCornerBase[j].Y := rCenterRobotY
                    + rLocalX * rSinTheta + rLocalY * rCosTheta;
                aQueue[nSlot].aCornerNow[j] := aQueue[nSlot].aCornerBase[j];
            END_FOR;
            nQueueCount := nQueueCount + 1;
            nAccepted := nAccepted + 1;
            nTailIndex := nTailIndex + 1;
            IF nTailIndex > 8 THEN nTailIndex := 1; END_IF;
            bPendingExposure := FALSE;
            nErrorCode := 0;
        END_IF;
    END_IF;

    // Tracking EVERY queued product each 10 ms using integrated encoder.
    // Future margin is only a conservative planning estimate, not a robot start permit.
    rForecastMotion_mm := 0.0;
    IF rConveyorSpeed_mm_s > 0.0 THEN
        rForecastMotion_mm := rConveyorSpeed_mm_s *
            (rMinCycleBudget_s + rFlyTime_s + rSyncTime_s);
    END_IF;
    FOR i := 1 TO 8 DO
        IF aQueue[i].bValid THEN
            aQueue[i].rTravel_mm := rEncoderTotalDist_mm -
                                      aQueue[i].rEncoderAtExposure_mm;
            aQueue[i].rCenterNowX_mm := aQueue[i].rCenterAtExposureX_mm +
                                        aQueue[i].rTravel_mm;
            aQueue[i].rCenterNowY_mm := aQueue[i].rCenterAtExposureY_mm;
            aQueue[i].bAllCornersInside := TRUE;
            aQueue[i].bForecastWindowOK := TRUE;
            FOR j := 1 TO 4 DO
                aQueue[i].aCornerNow[j].X := aQueue[i].aCornerBase[j].X +
                                            aQueue[i].rTravel_mm;
                aQueue[i].aCornerNow[j].Y := aQueue[i].aCornerBase[j].Y;
                IF (aQueue[i].aCornerNow[j].X < rXMin_mm)
                   OR (aQueue[i].aCornerNow[j].X > rXMax_mm)
                   OR (aQueue[i].aCornerNow[j].Y < rYMin_mm)
                   OR (aQueue[i].aCornerNow[j].Y > rYMax_mm) THEN
                    aQueue[i].bAllCornersInside := FALSE;
                END_IF;
                IF (aQueue[i].aCornerNow[j].X < rXMin_mm)
                   OR (aQueue[i].aCornerNow[j].X + rForecastMotion_mm > rXMax_mm)
                   OR (aQueue[i].aCornerNow[j].Y < rYMin_mm)
                   OR (aQueue[i].aCornerNow[j].Y > rYMax_mm) THEN
                    aQueue[i].bForecastWindowOK := FALSE;
                END_IF;
            END_FOR;
            IF aQueue[i].bAllCornersInside THEN
                aQueue[i].nState := 2; // all four corners geometrically in workspace
            ELSE
                aQueue[i].nState := 1;
            END_IF;
        END_IF;
    END_FOR;

    // Drop ONLY the oldest missed product; preserve FIFO order for later items.
    IF nQueueCount > 0 THEN
        bOut := TRUE;
        FOR j := 1 TO 4 DO
            IF aQueue[nHeadIndex].aCornerNow[j].X <= rXMax_mm THEN
                bOut := FALSE;
            END_IF;
        END_FOR;
        IF bOut THEN
            aQueue[nHeadIndex].bValid := FALSE;
            aQueue[nHeadIndex].nState := 0;
            nMissed := nMissed + 1;
            nQueueCount := nQueueCount - 1;
            nHeadIndex := nHeadIndex + 1;
            IF nHeadIndex > 8 THEN nHeadIndex := 1; END_IF;
        END_IF;
    END_IF;

    // Offline/manual simulation of completion only; never constitutes M1001 ACK.
    IF fbSimDoneEdge.Q AND (nQueueCount > 0) THEN
        IF aQueue[nHeadIndex].bAllCornersInside THEN
            aQueue[nHeadIndex].bValid := FALSE;
            aQueue[nHeadIndex].nState := 0;
            nSimCompleted := nSimCompleted + 1;
            nQueueCount := nQueueCount - 1;
            nHeadIndex := nHeadIndex + 1;
            IF nHeadIndex > 8 THEN nHeadIndex := 1; END_IF;
        ELSE
            nErrorCode := 116; // Simulation completion outside geometric window
        END_IF;
    END_IF;
END_IF;

// Presentation: active head is distinct from historical/legacy corner values.
bHeadValid := nQueueCount > 0;
bHeadAllInside := FALSE;
bHeadForecastOK := FALSE;
nHeadProductID := 0;
nHeadState := 0;
rHeadTravel_mm := 0.0;
rHeadToWorkStart_mm := 0.0;
rHeadCenterX_mm := 0.0;
rHeadCenterY_mm := 0.0;
FOR j := 1 TO 4 DO
    aHeadCornerNow[j].X := 0.0;
    aHeadCornerNow[j].Y := 0.0;
END_FOR;
IF bHeadValid THEN
    nHeadProductID := aQueue[nHeadIndex].nProductID;
    nHeadState := aQueue[nHeadIndex].nState;
    bHeadAllInside := aQueue[nHeadIndex].bAllCornersInside;
    bHeadForecastOK := aQueue[nHeadIndex].bForecastWindowOK;
    rHeadTravel_mm := aQueue[nHeadIndex].rTravel_mm;
    rHeadCenterX_mm := aQueue[nHeadIndex].rCenterNowX_mm;
    rHeadCenterY_mm := aQueue[nHeadIndex].rCenterNowY_mm;
    IF rHeadCenterX_mm < 0.0 THEN
        rHeadToWorkStart_mm := -rHeadCenterX_mm;
    END_IF;
    FOR j := 1 TO 4 DO
        aHeadCornerNow[j] := aQueue[nHeadIndex].aCornerNow[j];
    END_FOR;
END_IF;

END_FUNCTION_BLOCK

// ---- POUs/FB_XYTrackingManualAck.TcPOU
FUNCTION_BLOCK FB_XYTrackingManualAck
VAR_INPUT
    bExecute         : BOOL := FALSE;
    bPermit          : BOOL := FALSE; // OFF by default; user must approve spare PLC bit
    bAckBitAudited   : BOOL := FALSE; // Must be confirmed unused in PLC and HMI
    nAckAddress      : UDINT := 2100; // PROPOSED spare M, NOT M1001 or other motion bit
    bSafeToWriteXY   : BOOL := FALSE; // All other Publishers disabled; no robot motion
    bProductCaptured : BOOL;
    aCornerNow       : ARRAY[1..4] OF ST_Point2D;
    rConveyorSpeed   : LREAL;       // measured from encoder; may be zero for bench
    rFlyTime_s       : LREAL := 0.12;
    rXMax_mm         : LREAL := 180.0;
    rYMax_mm         : LREAL := 170.0;
    bAbort           : BOOL := FALSE;
END_VAR
VAR_IN_OUT
    stSession        : ST_MelsecSession;
END_VAR
VAR_OUTPUT
    bBusy            : BOOL;
    bDone            : BOOL; // DATA-ONLY: all four XY frames acknowledged MANUALLY
    bError           : BOOL;
    nErrorCode       : INT;
    nCommError       : UDINT;
    nState           : INT := 0;
    nVertex          : INT;
    nAckedVertices   : INT;
    bAckBitNow       : BOOL;
    nSentX           : DINT;
    nSentY           : DINT;
    nReadX           : DINT;
    nReadY           : DINT;
    nReadVertex      : UINT;
    bReadbackOK      : BOOL;
    bRestored        : BOOL;
END_VAR
VAR
    fbStart          : R_TRIG;
    fbWrite          : FB_MelsecWrite;
    fbRead           : FB_MelsecRead;
    tonWait          : TON;
    tonReview        : TON;
    aOriginalXY      : ARRAY[0..1] OF DINT;
    nOriginalIndex   : UINT;
    aWriteXY         : ARRAY[0..1] OF DINT;
    aReadXY          : ARRAY[0..1] OF DINT;
    nWriteIndex      : UINT;
    nReadIndex       : UINT;
    aStartAck        : ARRAY[0..1] OF BOOL; // M1000 M1001
    aRobotFlags      : ARRAY[0..3] OF BOOL; // M102..105
    nPlcState        : DINT;             // D200 D201
    bWriteReq        : BOOL;
    bReadReq         : BOOL;
    nWriteAddress    : UDINT;
    nWritePoints     : UINT;
    pWriteData       : PVOID;
    nWriteSize       : UDINT;
    eReadDevice      : E_MelsecDevice;
    nReadAddress     : UDINT;
    nReadPoints      : UINT;
    bReadBitMode     : BOOL;
    pReadData        : PVOID;
    nReadSize        : UDINT;
    rTargetX         : LREAL;
    rTargetY         : LREAL;
    bNeedOriginal    : BOOL;
    bRestoring       : BOOL;
END_VAR

// THIS IS NOT A ROBOT CYCLE. Never writes M1000, M1001, M105, Z or QD75.
// Operator toggles a separate AUDITED spare PLC bit M2100 for manual ack.
// M1001 is deliberately NOT used: the PLC owns it as true ROBOT DONE.
fbStart(CLK := bExecute);
tonWait(IN := bBusy AND NOT bRestoring AND (nState >= 10) AND
            (nState <= 25), PT := T#25S);
tonReview(IN := (nState = 23) OR (nState = 24), PT := T#2S);
bWriteReq := FALSE;
bReadReq := FALSE;

IF (nState <> 0) AND (nState <> 99) AND
   (NOT bPermit OR NOT bAckBitAudited OR NOT bSafeToWriteXY OR
    bAbort OR NOT stSession.bConnected OR NOT bProductCaptured) THEN
    bError := TRUE;
    nErrorCode := 901;
    nState := 99;
END_IF;

CASE nState OF
    0:
        bBusy := FALSE;
        IF fbStart.Q THEN
            bDone := FALSE; bError := FALSE; bRestored := FALSE;
            nErrorCode := 0; nCommError := 0;
            nAckedVertices := 0; nVertex := 0;
            bReadbackOK := FALSE;
            IF NOT bPermit OR NOT bAckBitAudited OR NOT bSafeToWriteXY OR
               NOT bProductCaptured OR bAbort OR NOT stSession.bConnected OR
               stSession.bBusy OR (nAckAddress < 2000) OR (nAckAddress > 8191) THEN
                bError := TRUE; nErrorCode := 901;
            ELSE
                bBusy := TRUE; bNeedOriginal := TRUE;
                bRestoring := FALSE;
                nVertex := 1; nState := 1;
            END_IF;
        END_IF;

    1: // Motion handshake must stay LOW
        eReadDevice := DEV_M; nReadAddress := 1000; nReadPoints := 2;
        bReadBitMode := TRUE;
        pReadData := ADR(aStartAck); nReadSize := SIZEOF(aStartAck);
        bReadReq := TRUE; nState := 2;

    2:
        IF fbRead.bDone THEN
            IF aStartAck[0] OR aStartAck[1] THEN
                bError := TRUE; nErrorCode := 902; nState := 99;
            ELSE
                nState := 3;
            END_IF;
        ELSIF fbRead.bError THEN
            bError := TRUE; nErrorCode := 910; nCommError := fbRead.nErrorID; nState := 99;
        END_IF;

    3:
        eReadDevice := DEV_M; nReadAddress := 102; nReadPoints := 4;
        bReadBitMode := TRUE;
        pReadData := ADR(aRobotFlags); nReadSize := SIZEOF(aRobotFlags);
        bReadReq := TRUE; nState := 4;

    4:
        IF fbRead.bDone THEN
            IF aRobotFlags[0] OR aRobotFlags[1] OR aRobotFlags[2] OR aRobotFlags[3] THEN
                bError := TRUE; nErrorCode := 903; nState := 99;
            ELSE
                nState := 5;
            END_IF;
        ELSIF fbRead.bError THEN
            bError := TRUE; nErrorCode := 911; nCommError := fbRead.nErrorID; nState := 99;
        END_IF;

    5:
        eReadDevice := DEV_D; nReadAddress := 200; nReadPoints := 2;
        bReadBitMode := FALSE;
        pReadData := ADR(nPlcState); nReadSize := SIZEOF(nPlcState);
        bReadReq := TRUE; nState := 6;

    6:
        IF fbRead.bDone THEN
            IF nPlcState <> 0 THEN
                bError := TRUE; nErrorCode := 904; nState := 99;
            ELSE
                nState := 7;
            END_IF;
        ELSIF fbRead.bError THEN
            bError := TRUE; nErrorCode := 912; nCommError := fbRead.nErrorID; nState := 99;
        END_IF;

    7: // Require manual ACK LOW before a new vertex
        eReadDevice := DEV_M; nReadAddress := nAckAddress; nReadPoints := 1;
        bReadBitMode := TRUE;
        pReadData := ADR(bAckBitNow); nReadSize := SIZEOF(bAckBitNow);
        bReadReq := TRUE; nState := 8;

    8:
        IF fbRead.bDone THEN
            IF bAckBitNow THEN
                bError := TRUE; nErrorCode := 905; nState := 99;
            ELSIF bNeedOriginal THEN
                nState := 30;
            ELSIF bRestoring THEN
                nState := 40;
            ELSE
                nState := 10;
            END_IF;
        ELSIF fbRead.bError THEN
            bError := TRUE; nErrorCode := 913; nCommError := fbRead.nErrorID; nState := 99;
        END_IF;

    30: // Save X/Y and index to restore after four acknowledgements
        eReadDevice := DEV_D; nReadAddress := 100; nReadPoints := 4;
        bReadBitMode := FALSE;
        pReadData := ADR(aOriginalXY); nReadSize := SIZEOF(aOriginalXY);
        bReadReq := TRUE; nState := 31;

    31:
        IF fbRead.bDone THEN nState := 32;
        ELSIF fbRead.bError THEN
            bError := TRUE; nErrorCode := 914; nCommError := fbRead.nErrorID; nState := 99;
        END_IF;

    32:
        eReadDevice := DEV_D; nReadAddress := 114; nReadPoints := 1;
        bReadBitMode := FALSE;
        pReadData := ADR(nOriginalIndex); nReadSize := SIZEOF(nOriginalIndex);
        bReadReq := TRUE; nState := 33;

    33:
        IF fbRead.bDone THEN
            bNeedOriginal := FALSE; nState := 10;
        ELSIF fbRead.bError THEN
            bError := TRUE; nErrorCode := 915; nCommError := fbRead.nErrorID; nState := 99;
        END_IF;

    10: // Live computation directly before EACH vertex write
        rTargetX := aCornerNow[nVertex].X + rConveyorSpeed * rFlyTime_s;
        rTargetY := aCornerNow[nVertex].Y;
        IF (ABS(rConveyorSpeed) > 1000.0) OR
            (rTargetY < 0.0) OR (rTargetY > rYMax_mm) OR
            (rTargetX > rXMax_mm) THEN
            bError := TRUE; nErrorCode := 906; nState := 99;
        ELSIF rTargetX < 0.0 THEN
            // Camera is upstream: WAIT for tracked vertex to reach workspace
            IF tonWait.Q THEN
                bError := TRUE; nErrorCode := 907; nState := 99;
            END_IF;
        ELSE
            nSentX := LREAL_TO_DINT(rTargetX * 10000.0);
            nSentY := LREAL_TO_DINT(rTargetY * 10000.0);
            aWriteXY[0] := nSentX;
            aWriteXY[1] := nSentY;
            nWriteIndex := INT_TO_UINT(nVertex);
            nWriteAddress := 100; nWritePoints := 4;
            pWriteData := ADR(aWriteXY); nWriteSize := SIZEOF(aWriteXY);
            bReadbackOK := FALSE;
            bWriteReq := TRUE; nState := 11;
        END_IF;

    11:
        IF fbWrite.bDone THEN nState := 12;
        ELSIF fbWrite.bError THEN
            bError := TRUE; nErrorCode := 916; nCommError := fbWrite.nErrorID; nState := 99;
        END_IF;

    12:
        nWriteAddress := 114; nWritePoints := 1;
        pWriteData := ADR(nWriteIndex); nWriteSize := SIZEOF(nWriteIndex);
        bWriteReq := TRUE; nState := 13;

    13:
        IF fbWrite.bDone THEN nState := 14;
        ELSIF fbWrite.bError THEN
            bError := TRUE; nErrorCode := 917; nCommError := fbWrite.nErrorID; nState := 99;
        END_IF;

    14:
        eReadDevice := DEV_D; nReadAddress := 100; nReadPoints := 4;
        bReadBitMode := FALSE;
        pReadData := ADR(aReadXY); nReadSize := SIZEOF(aReadXY);
        bReadReq := TRUE; nState := 15;

    15:
        IF fbRead.bDone THEN nState := 16;
        ELSIF fbRead.bError THEN
            bError := TRUE; nErrorCode := 918; nCommError := fbRead.nErrorID; nState := 99;
        END_IF;

    16:
        eReadDevice := DEV_D; nReadAddress := 114; nReadPoints := 1;
        bReadBitMode := FALSE;
        pReadData := ADR(nReadIndex); nReadSize := SIZEOF(nReadIndex);
        bReadReq := TRUE; nState := 17;

    17:
        IF fbRead.bDone THEN
            nReadX := aReadXY[0]; nReadY := aReadXY[1]; nReadVertex := nReadIndex;
            bReadbackOK := (nReadX = nSentX) AND (nReadY = nSentY)
                           AND (nReadVertex = nWriteIndex);
            IF bReadbackOK THEN nState := 20;
            ELSE bError := TRUE; nErrorCode := 919; nState := 99;
            END_IF;
        ELSIF fbRead.bError THEN
            bError := TRUE; nErrorCode := 920; nCommError := fbRead.nErrorID; nState := 99;
        END_IF;

    20: // Wait for human acknowledgement at separately reserved PLC M bit
        IF (aCornerNow[nVertex].X > rXMax_mm) OR tonWait.Q THEN
            bError := TRUE; nErrorCode := 921; nState := 99;
        ELSE
            eReadDevice := DEV_M; nReadAddress := nAckAddress; nReadPoints := 1;
            bReadBitMode := TRUE;
            pReadData := ADR(bAckBitNow); nReadSize := SIZEOF(bAckBitNow);
            bReadReq := TRUE; nState := 21;
        END_IF;

    21:
        IF fbRead.bDone THEN
            IF bAckBitNow THEN
                nAckedVertices := nAckedVertices + 1;
                nState := 23;
            ELSE
                nState := 20;
            END_IF;
        ELSIF fbRead.bError THEN
            bError := TRUE; nErrorCode := 922; nCommError := fbRead.nErrorID; nState := 99;
        END_IF;

    23: // Show acknowledged point for >=2 s only when conveyor is stationary
        IF (ABS(rConveyorSpeed) > 1.0) OR tonReview.Q THEN
            nState := 24;
        END_IF;

    24: // Operator must clear ACK before TwinCAT computes next tracked corner
        IF (aCornerNow[nVertex].X > rXMax_mm) OR tonWait.Q THEN
            bError := TRUE; nErrorCode := 923; nState := 99;
        ELSE
            eReadDevice := DEV_M; nReadAddress := nAckAddress; nReadPoints := 1;
            bReadBitMode := TRUE;
            pReadData := ADR(bAckBitNow); nReadSize := SIZEOF(bAckBitNow);
            bReadReq := TRUE; nState := 25;
        END_IF;

    25:
        IF fbRead.bDone THEN
            IF NOT bAckBitNow THEN
                IF nVertex >= 4 THEN
                    bRestoring := TRUE; nState := 1;
                ELSE
                    nVertex := nVertex + 1; nState := 1;
                END_IF;
            ELSE
                nState := 24;
            END_IF;
        ELSIF fbRead.bError THEN
            bError := TRUE; nErrorCode := 924; nCommError := fbRead.nErrorID; nState := 99;
        END_IF;

    40:
        nWriteAddress := 100; nWritePoints := 4;
        pWriteData := ADR(aOriginalXY); nWriteSize := SIZEOF(aOriginalXY);
        bWriteReq := TRUE; nState := 41;
    41:
        IF fbWrite.bDone THEN nState := 42;
        ELSIF fbWrite.bError THEN
            bError := TRUE; nErrorCode := 925; nCommError := fbWrite.nErrorID; nState := 99;
        END_IF;
    42:
        nWriteAddress := 114; nWritePoints := 1;
        pWriteData := ADR(nOriginalIndex); nWriteSize := SIZEOF(nOriginalIndex);
        bWriteReq := TRUE; nState := 43;
    43:
        IF fbWrite.bDone THEN nState := 44;
        ELSIF fbWrite.bError THEN
            bError := TRUE; nErrorCode := 926; nCommError := fbWrite.nErrorID; nState := 99;
        END_IF;
    44:
        eReadDevice := DEV_D; nReadAddress := 100; nReadPoints := 4;
        bReadBitMode := FALSE;
        pReadData := ADR(aReadXY); nReadSize := SIZEOF(aReadXY);
        bReadReq := TRUE; nState := 45;
    45:
        IF fbRead.bDone THEN nState := 46;
        ELSIF fbRead.bError THEN
            bError := TRUE; nErrorCode := 927; nCommError := fbRead.nErrorID; nState := 99;
        END_IF;
    46:
        eReadDevice := DEV_D; nReadAddress := 114; nReadPoints := 1;
        bReadBitMode := FALSE;
        pReadData := ADR(nReadIndex); nReadSize := SIZEOF(nReadIndex);
        bReadReq := TRUE; nState := 47;
    47:
        IF fbRead.bDone THEN
            bRestored := (aReadXY[0] = aOriginalXY[0]) AND
                          (aReadXY[1] = aOriginalXY[1]) AND
                          (nReadIndex = nOriginalIndex);
            IF bRestored THEN
                bBusy := FALSE; bDone := TRUE; nState := 0;
            ELSE
                bError := TRUE; nErrorCode := 928; nState := 99;
            END_IF;
        ELSIF fbRead.bError THEN
            bError := TRUE; nErrorCode := 929; nCommError := fbRead.nErrorID; nState := 99;
        END_IF;

    99: // Fail closed, no robot command
        bBusy := FALSE; bDone := FALSE;
        IF NOT bExecute AND NOT bPermit AND NOT fbRead.bBusy AND NOT fbWrite.bBusy THEN
            nState := 0;
        END_IF;
END_CASE;

// MC 3E Client sends exactly these XY-only word regions; no M write possible.
fbWrite(stSession := stSession, bExecute := bWriteReq,
        eDevice := DEV_D, nStartAddr := nWriteAddress,
        nPoints := nWritePoints, bBitAccess := FALSE,
        pData := pWriteData, nDataSize := nWriteSize);
fbRead(stSession := stSession, bExecute := bReadReq,
       eDevice := eReadDevice, nStartAddr := nReadAddress,
       nPoints := nReadPoints, bBitAccess := bReadBitMode,
       pData := pReadData, nDataSize := nReadSize);

END_FUNCTION_BLOCK

// ---- POUs/FB_MelsecEchoVerify.TcPOU
FUNCTION_BLOCK FB_MelsecEchoVerify
VAR_INPUT
    bExecute                : BOOL;          // Rising edge starts one write/read/restore cycle
    bEnable                 : BOOL := FALSE; // OFF by default
    bAddressVerifiedUnused  : BOOL := FALSE; // Operator approved address in real PLC/HMI
    bMachineSafe            : BOOL := FALSE; // Operator confirmed safe machine state
    bBitDevice              : BOOL := FALSE; // FALSE -> D word, TRUE -> M bit
    nAddress                : UDINT := 0;    // D>=3000 or M>=2000; still requires approval
    wTestValue              : WORD := 16#A55A;
    bTestValue              : BOOL := TRUE;
END_VAR
VAR_IN_OUT
    stSession               : ST_MelsecSession;
END_VAR
VAR_OUTPUT
    bBusy                   : BOOL;
    bDone                   : BOOL;          // Complete after restore verification
    bError                  : BOOL;
    bMatch                  : BOOL;          // Readback equals test value
    bRestored               : BOOL;          // PLC reply confirms original value
    bRestoreUncertain       : BOOL;          // A write may have happened before error
    nErrorID                : UDINT;
    nState                  : INT;
    wOriginal               : WORD;
    wReadBack               : WORD;
    bOriginal               : BOOL;
    bReadBack               : BOOL;
END_VAR
VAR
    fbStart                 : R_TRIG;
    fbRead                  : FB_MelsecRead;
    fbWrite                 : FB_MelsecWrite;
    tonCycle                : TON;
    bReadReq                : BOOL;
    bWriteReq               : BOOL;
    bIsBit                  : BOOL;
    nSafeAddress            : UDINT;
    eSafeDevice             : E_MelsecDevice;
    nBufferSize             : UDINT;
    pReadBuffer             : PVOID;
    pWriteBuffer            : PVOID;
    wPayload                : WORD;
    bPayload                : BOOL;
    wCurrent                : WORD;
    bCurrent                : BOOL;
    wExpected               : WORD;
    bExpected               : BOOL;
END_VAR

fbStart(CLK := bExecute);
tonCycle(IN := bBusy, PT := T#25S);
bReadReq := FALSE;
bWriteReq := FALSE;

// Never start automatically: all three authorizations and an explicit edge are required.
IF (nState = 0) AND fbStart.Q THEN
    bDone := FALSE;
    bError := FALSE;
    bMatch := FALSE;
    bRestored := FALSE;
    bRestoreUncertain := FALSE;
    nErrorID := 0;
    IF NOT bEnable OR NOT bAddressVerifiedUnused OR NOT bMachineSafe THEN
        bError := TRUE; nErrorID := 16#E701; // Not authorized
    ELSIF NOT stSession.bConnected OR stSession.bBusy THEN
        bError := TRUE; nErrorID := 16#E702; // No free connected session
    ELSIF (bBitDevice AND ((nAddress < 2000) OR (nAddress > 8191)))
       OR ((NOT bBitDevice) AND ((nAddress < 3000) OR (nAddress > 7999))) THEN
        bError := TRUE; nErrorID := 16#E703; // Reserve low ranges for machine
    ELSE
        bIsBit := bBitDevice;
        nSafeAddress := nAddress;
        wExpected := wTestValue;
        bExpected := bTestValue;
        IF bIsBit THEN
            eSafeDevice := DEV_M;
            nBufferSize := SIZEOF(bCurrent);
            pReadBuffer := ADR(bCurrent);
            pWriteBuffer := ADR(bPayload);
        ELSE
            eSafeDevice := DEV_D;
            nBufferSize := SIZEOF(wCurrent);
            pReadBuffer := ADR(wCurrent);
            pWriteBuffer := ADR(wPayload);
        END_IF;
        bBusy := TRUE;
        nState := 10;
    END_IF;
END_IF;

IF bBusy AND tonCycle.Q THEN
    bError := TRUE;
    nErrorID := 16#E704; // Complete transaction did not finish in time
    bBusy := FALSE;
    nState := 0;
END_IF;

// One request at a time, with a scan gap between consecutive R_TRIG requests.
CASE nState OF
    10: // Read original before any write
        bReadReq := TRUE;
        nState := 11;
    11:
        IF fbRead.bError THEN
            bError := TRUE; nErrorID := fbRead.nErrorID;
            bBusy := FALSE; nState := 0;
        ELSIF fbRead.bDone THEN
            IF bIsBit THEN
                bOriginal := bCurrent;
                IF bOriginal = bExpected THEN
                    bError := TRUE; nErrorID := 16#E707; // Must change the bit to prove WRITE
                    bBusy := FALSE; nState := 0;
                ELSE nState := 20; END_IF;
            ELSE
                wOriginal := wCurrent;
                IF wOriginal = wExpected THEN
                    bError := TRUE; nErrorID := 16#E707; // Must change the word to prove WRITE
                    bBusy := FALSE; nState := 0;
                ELSE nState := 20; END_IF;
            END_IF;
        END_IF;

    20: // Write one approved device only
        IF bIsBit THEN bPayload := bExpected;
        ELSE wPayload := wExpected; END_IF;
        bRestoreUncertain := TRUE; // From now on, a failed call might have modified PLC
        bWriteReq := TRUE;
        nState := 21;
    21:
        IF fbWrite.bError THEN
            bError := TRUE; nErrorID := fbWrite.nErrorID;
            bBusy := FALSE; nState := 0;
        ELSIF fbWrite.bDone THEN
            nState := 30;
        END_IF;

    30: // Read exact same address
        bReadReq := TRUE;
        nState := 31;
    31:
        IF fbRead.bError THEN
            bError := TRUE; nErrorID := fbRead.nErrorID;
            bBusy := FALSE; nState := 0;
        ELSIF fbRead.bDone THEN
            IF bIsBit THEN
                bReadBack := bCurrent;
                bMatch := (bReadBack = bExpected);
            ELSE
                wReadBack := wCurrent;
                bMatch := (wReadBack = wExpected);
            END_IF;
            // Restore even after a mismatch, never leave the test value in the PLC.
            nState := 40;
        END_IF;

    40: // Restore original
        IF bIsBit THEN bPayload := bOriginal;
        ELSE wPayload := wOriginal; END_IF;
        bWriteReq := TRUE;
        nState := 41;
    41:
        IF fbWrite.bError THEN
            bError := TRUE; nErrorID := fbWrite.nErrorID;
            bBusy := FALSE; nState := 0;
        ELSIF fbWrite.bDone THEN
            nState := 50;
        END_IF;

    50: // Verify restoration from PLC
        bReadReq := TRUE;
        nState := 51;
    51:
        IF fbRead.bError THEN
            bError := TRUE; nErrorID := fbRead.nErrorID;
            bBusy := FALSE; nState := 0;
        ELSIF fbRead.bDone THEN
            IF bIsBit THEN bRestored := (bCurrent = bOriginal);
            ELSE bRestored := (wCurrent = wOriginal); END_IF;
            bRestoreUncertain := NOT bRestored;
            IF NOT bRestored THEN
                bError := TRUE; nErrorID := 16#E706; // Restore readback differs
            ELSIF NOT bMatch THEN
                bError := TRUE; nErrorID := 16#E705; // Test readback differs
            ELSE
                bDone := TRUE;
            END_IF;
            bBusy := FALSE;
            nState := 0;
        END_IF;
END_CASE;

// Exclusive access through ST_MelsecSession.bBusy in the existing MC FBs.
fbRead(
    stSession := stSession, bExecute := bReadReq,
    eDevice := eSafeDevice, nStartAddr := nSafeAddress,
    nPoints := 1, bBitAccess := bIsBit,
    pData := pReadBuffer, nDataSize := nBufferSize
);
fbWrite(
    stSession := stSession, bExecute := bWriteReq,
    eDevice := eSafeDevice, nStartAddr := nSafeAddress,
    nPoints := 1, bBitAccess := bIsBit,
    pData := pWriteBuffer, nDataSize := nBufferSize
);

END_FUNCTION_BLOCK
